FUNCTION_BLOCK F_NOT_BOOL_INIT (* standard boolean NOT function with INIT - wrapt F_NOT_BOOL, reicht INIT direkt auf INITO durch *)
  (* Standard: 61131-3; Classification: standard boolean function; Description: Copyright (c) 2011 TU Wien ACIN, HR Agrartechnik GmbH This program and the accompanying materials are made available under the terms of the Eclipse Public License 2.0 which is available at https://www.eclipse.org/legal/epl-2.0/ SPDX-License-Identifier: EPL-2.0 *)
  (* Version 3.1, 2026-10-11, Franz Höpfinger, Meisterschulen am Ostbahnhof, Interne Umsetzung wrapt jetzt den paketinternen F_NOT_BOOL statt iec61131::bitwiseOperators::F_NOT - damit entfaellt die letzte iec61131-3-Abhaengigkeit dieses Pakets. Instanzname F_NOT auf Negate umbenannt. Organization-Attribut ergaenzt (XSD-Pflichtfeld). *)
  (* Version 3.0, 2025-04-14, Patrick Aigner, Eclipse 4diac, changed package *)
  (* Version 1.0, 2011-06-21, Monika Wenger, TU Wien ACIN, initial API and implementation and/or initial documentation *)
  PACKAGE iec61131::booleanOperators;
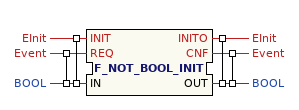
  EVENT_INPUT
    INIT : EInit WITH IN; (* Initialization Request *)
    REQ WITH IN; (* Service Request *)
  END_EVENT
  EVENT_OUTPUT
    INITO : EInit WITH OUT; (* Initialization Confirm *)
    CNF WITH OUT; (* Confirmation of Requested Service *)
  END_EVENT
  VAR_INPUT
    IN : BOOL; (* Input *)
  END_VAR
  VAR_OUTPUT
    OUT : BOOL; (* Output *)
  END_VAR
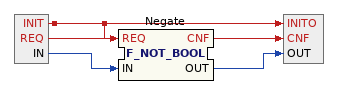
  FBS
    Negate : iec61131::booleanOperators::F_NOT_BOOL;
  END_FBS
  EVENT_CONNECTIONS
    REQ TO Negate.REQ;
    Negate.CNF TO CNF;
    INIT TO INITO;
    INIT TO Negate.REQ;
  END_CONNECTIONS
  DATA_CONNECTIONS
    IN TO Negate.IN;
    Negate.OUT TO OUT;
  END_CONNECTIONS
END_FUNCTION_BLOCK
